(* Communication structure from plc to drive *)

TYPE ST_PLCTOSEWMOVIEDRIVEBCIA402 :
STRUCT
	wPO1ControlWord			:WORD;
END_STRUCT
END_TYPE

(* stored: Version 1.1.0.1, ProductVersion 3.1.4024.15
   DUT ST_PLCTOSEWMOVIEDRIVEBCIA402: Id {2a9394fa-ac09-4857-9994-76e9bebb2c5c} *)
